{attribute 'qualified_only'}
VAR_GLOBAL
	RedLED 			  AT %Q*: BOOL;
	GreenLED 		  AT %Q*: BOOL;
	BlueLED			  AT %Q*: BOOL;
	b_MotorCooling			  AT %Q*: BOOL;
	    // I/O module state — Python can read inputs and write output setpoints
    // ADS symbol: GVL_IO.stIO
    stIO            : ST_IOData;

END_VAR

(* stored: Version 1.1.0.1, ProductVersion 3.1.4026.18
   GVL GVL_IO: Id {480a6fec-3a96-474a-a55b-a1de807d8f3f} *)
